Fanuc KAREL source: KT00163.KL

PROGRAM KT00163
%NOLOCKGROUP
VAR
  I1: INTEGER
  R2: REAL
  OUT: INTEGER
BEGIN
  I1 = 2
    R2 = 3.0
  OUT = I1 MOD R2
END KT00163
